{region 'Documentation'}
(*!
<summary>Check that IN is outside the inclusive StartTime..EndTime interval.</summary>
<description>

StartTime &gt; EndTime reports Error during active evaluation; equal bounds are
valid.

</description>
*)
{endregion}
FUNCTION_BLOCK AssertNotInTimespan_Time EXTENDS AssertionBase
VAR_INPUT
    IN : TIME; //! Actual value checked or observed by this Assertion.
    StartTime : TIME; //! Inclusive start of the time span; must not exceed EndTime.
    EndTime : TIME; //! Inclusive end of the time span; must not precede StartTime.
END_VAR

SUPER^();

{region 'Documentation'}
(*!
<summary>Evaluate the typed duration relation and report higher-priority errors first.</summary>
*)
{endregion}
METHOD PROTECTED Assert
VAR
    Message : STRING(GVL_Constants.MessageLength);
    StartTimeText : STRING(GVL_Constants.AssertionValueLength);
    EndTimeText : STRING(GVL_Constants.AssertionValueLength);
    ActualText : STRING(GVL_Constants.AssertionValueLength);
END_VAR
IF NOT EvaluationActive THEN
    RETURN;
END_IF;

IF Result = E_Result.Error THEN
    RETURN;
END_IF;

IF StartTime > EndTime THEN
    StartTimeText := TIME_TO_STRING(StartTime);
    EndTimeText := TIME_TO_STRING(EndTime);
    Message := CONCAT('Assertion error: start time exceeds end time. StartTime = ',
        StartTimeText);
    Message := CONCAT(Message, ', EndTime = ');
    Message := CONCAT(Message, EndTimeText);
    Message := CONCAT(Message, '.');
    Error(Message := Message);
    RETURN;
END_IF;

IF Result = E_Result.Failed THEN
    RETURN;
END_IF;

IF (IN >= StartTime) AND (IN <= EndTime) THEN
    StartTimeText := TIME_TO_STRING(StartTime);
    EndTimeText := TIME_TO_STRING(EndTime);
    ActualText := TIME_TO_STRING(IN);
    Message := CONCAT('Assertion failed: value is inside forbidden timespan. StartTime = ',
        StartTimeText);
    Message := CONCAT(Message, ', EndTime = ');
    Message := CONCAT(Message, EndTimeText);
    Message := CONCAT(Message, ', Actual = ');
    Message := CONCAT(Message, ActualText);
    Message := CONCAT(Message, '.');
    Fail(Message := Message);
    RETURN;
END_IF;

Pass();
END_METHOD

END_FUNCTION_BLOCK

(* stored: Version 1.1.0.1
   POU AssertNotInTimespan_Time: Id {20ed8b88-5513-4863-93f9-afb67215b089}, SpecialFunc None
   Folder Internal: Id {51b3ee6e-0588-4819-bbe6-06b2424ae8f2}
   Method Assert: Id {14c3f24a-9e19-448d-9131-6d4f3585d2b8} *)
